// TIA Portal V21 export
FUNCTION_BLOCK "FB_BackwashGraph"   // FB120, GRAPH
TITLE = Промывка фильтра (GRAPH)
{ S7_Optimized_Access := 'TRUE' }
AUTHOR : WTP2
FAMILY : Filters
VERSION : 0.1
// Промывка скорого фильтра (GRAPH S7-1500), шаги S1–S6. S1 Idle (начальный): N xReady.
// T1 Start: xStart. S2 Drain: N xDrainValve, S xWashActive, событие S1 — iWashCount + 1;
// контроль xValveFault держит шаг до квитирования ACK_EF (ERR_FLT = 1). После S2 альтернатива:
// T2 LongWash (xLevelLow AND NOT xShortWash) — параллельно S3 Air (N xBlower, D xAirValve 2 с)
// и S4 Rinse (NC xWashPump, блокировка xPumpOk), синхронизация T4 AirDone: Air.T >= 10 с;
// T3 ShortWash (xLevelLow AND xShortWash) — S5 QuickRinse (N xWashPump), T5 QuickDone: xLevelHigh.
// S6 Refill: N xInletValve, R xWashActive; T6 Full: xLevelHigh — прыжок к S1. Постоперация:
// xValvesBusy := xDrainValve OR xInletValve. INIT_SQ — начальное состояние, OFF_SQ — шаги выключены.
// stored: AutoNumber false, SetENOAutomatically false
   VAR_INPUT
      OFF_SQ : Bool;   // Выключить последовательность
      INIT_SQ : Bool;   // Начальное состояние
      ACK_EF : Bool;   // Квитирование ошибок контроля
      xStart : Bool;   // Пуск промывки
      xLevelLow : Bool;   // Уровень ниже сливного
      xLevelHigh : Bool;   // Фильтр заполнен
      xShortWash : Bool;   // Короткая промывка (без продувки)
      xPumpOk : Bool := TRUE;   // Насос промывки исправен
      xValveFault : Bool;   // Неисправность сливной задвижки
   END_VAR
   VAR_OUTPUT
      ERR_FLT : Bool;   // Ошибка контроля (до квитирования)
      xReady : Bool;   // Готов к промывке
      xDrainValve : Bool;   // Сливная задвижка
      xBlower : Bool;   // Воздуходувка
      xAirValve : Bool;   // Задвижка воздуха
      xWashPump : Bool;   // Насос промывки
      xInletValve : Bool;   // Задвижка подачи
      xWashActive : Bool;   // Промывка идёт
      xValvesBusy : Bool;   // Задвижки в работе
      iWashCount : Int;   // Число промывок
   END_VAR
BEGIN
// Промывка фильтра
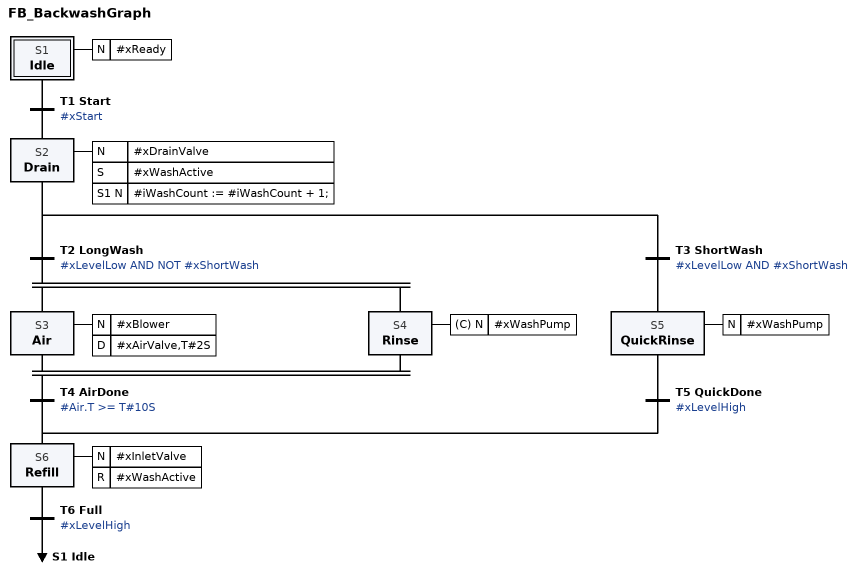
   // sequencer 1
   INITIAL_STEP Idle:   // S1
              N    #xReady
   END_STEP
   TRANSITION Start FROM Idle TO Drain   // T1
      := #xStart;
   END_TRANSITION
   STEP Drain:   // S2
      supervision V := #xValveFault;
              N    #xDrainValve
              S    #xWashActive
          S1  N    #iWashCount := #iWashCount + 1;
   END_STEP
   TRANSITION LongWash FROM Drain TO (Air, Rinse)   // T2
      := #xLevelLow AND NOT #xShortWash;
   END_TRANSITION
   TRANSITION ShortWash FROM Drain TO QuickRinse   // T3
      := #xLevelLow AND #xShortWash;
   END_TRANSITION
   STEP Air:   // S3
              N    #xBlower
              D    #xAirValve,T#2S
   END_STEP
   STEP Rinse:   // S4
      interlock C := #xPumpOk;
      (C)     N    #xWashPump
   END_STEP
   TRANSITION AirDone FROM (Air, Rinse) TO Refill   // T4
      := #Air.T >= T#10S;
   END_TRANSITION
   STEP QuickRinse:   // S5
              N    #xWashPump
   END_STEP
   TRANSITION QuickDone FROM QuickRinse TO Refill   // T5
      := #xLevelHigh;
   END_TRANSITION
   STEP Refill:   // S6
              N    #xInletValve
              R    #xWashActive
   END_STEP
   TRANSITION Full FROM Refill TO Idle   // T6, jump
      := #xLevelHigh;
   END_TRANSITION

   // permanent post-instructions
   NETWORK 1
      #xValvesBusy := #xDrainValve OR #xInletValve;
END_FUNCTION_BLOCK
